(* IEC 61131-3 sources: llm-plc-st-eval/data/processed_definitivo/gpt-4o-2024-08-06/C4/zero_shot, 3 files *)

(* ---- ejec_1.st ---- *)
FUNCTION_BLOCK FB_D
VAR_INPUT
    demanda : BOOL;  // Entrada que indica si hay demanda para activar las bombas.
    falla1 : BOOL;   // Entrada que indica si la bomba1 tiene una falla.
    falla2 : BOOL;   // Entrada que indica si la bomba2 tiene una falla.
END_VAR
VAR_OUTPUT
    bomba1 : BOOL;   // Salida que controla el estado de la bomba1 (activa/inactiva).
    bomba2 : BOOL;   // Salida que controla el estado de la bomba2 (activa/inactiva).
    almFalla : BOOL; // Salida que indica si hay una alarma de falla en la bomba activa.
END_VAR
VAR
    turno : BOOL;    // Variable interna que determina cuál bomba debe activarse.
    fDem : R_TRIG;   // Detector de flanco ascendente para la señal de demanda.
END_VAR

// Detecta el flanco ascendente de la señal de demanda.
fDem(CLK := demanda);

// Si se detecta un flanco ascendente en la demanda, alterna el turno.
IF fDem.Q THEN
    turno := NOT turno;
END_IF

// Si hay demanda, decide qué bomba activar según el turno y el estado de fallas.
IF demanda THEN
    IF turno THEN
        // Si es el turno de la bomba1, actívala si no hay falla.
        bomba1 := NOT falla1;
        // Activa la bomba2 solo si la bomba1 falla y la bomba2 no tiene falla.
        bomba2 := falla1 AND NOT falla2;
        // Genera alarma si la bomba1 tiene falla.
        almFalla := falla1;
    ELSE
        // Si es el turno de la bomba2, actívala si no hay falla.
        bomba2 := NOT falla2;
        // Activa la bomba1 solo si la bomba2 falla y la bomba1 no tiene falla.
        bomba1 := falla2 AND NOT falla1;
        // Genera alarma si la bomba2 tiene falla.
        almFalla := falla2;
    END_IF
ELSE
    // Si no hay demanda, ambas bombas están inactivas y no hay alarma.
    bomba1 := FALSE;
    bomba2 := FALSE;
    almFalla := FALSE;
END_IF
END_FUNCTION_BLOCK

(* ---- ejec_2.st ---- *)
FUNCTION_BLOCK FB_D
VAR_INPUT
    demanda : BOOL; // Entrada que indica si hay demanda de bombeo
    falla1 : BOOL;  // Entrada que indica si la bomba 1 ha fallado
    falla2 : BOOL;  // Entrada que indica si la bomba 2 ha fallado
END_VAR
VAR_OUTPUT
    bomba1 : BOOL;  // Salida que controla el estado de la bomba 1
    bomba2 : BOOL;  // Salida que controla el estado de la bomba 2
    almFalla : BOOL; // Salida que indica si hay una alarma de falla
END_VAR
VAR
    turno : BOOL;   // Variable interna para alternar el uso de las bombas
    fDem : R_TRIG;  // Detector de flanco ascendente para la señal de demanda
END_VAR

// Detecta un flanco ascendente en la señal de demanda
fDem(CLK := demanda);

// Si se detecta un flanco ascendente en la demanda, alterna el turno
IF fDem.Q THEN
    turno := NOT turno;
END_IF

// Si hay demanda de bombeo
IF demanda THEN
    // Si es el turno de la bomba 1
    IF turno THEN
        bomba1 := NOT falla1; // Activa la bomba 1 si no hay falla
        bomba2 := falla1 AND NOT falla2; // Activa la bomba 2 si la bomba 1 falla y la bomba 2 no
        almFalla := falla1; // Activa la alarma si la bomba 1 falla
    ELSE
        // Si es el turno de la bomba 2
        bomba2 := NOT falla2; // Activa la bomba 2 si no hay falla
        bomba1 := falla2 AND NOT falla1; // Activa la bomba 1 si la bomba 2 falla y la bomba 1 no
        almFalla := falla2; // Activa la alarma si la bomba 2 falla
    END_IF
ELSE
    // Si no hay demanda, apaga ambas bombas y resetea la alarma
    bomba1 := FALSE;
    bomba2 := FALSE;
    almFalla := FALSE;
END_IF
END_FUNCTION_BLOCK

(* ---- ejec_3.st ---- *)
FUNCTION_BLOCK FB_D
VAR_INPUT
    demanda : BOOL;  // Entrada que indica si hay demanda de bombeo.
    falla1 : BOOL;   // Entrada que indica si la bomba1 está en estado de falla.
    falla2 : BOOL;   // Entrada que indica si la bomba2 está en estado de falla.
END_VAR
VAR_OUTPUT
    bomba1 : BOOL;   // Salida que controla el estado de la bomba1.
    bomba2 : BOOL;   // Salida que controla el estado de la bomba2.
    almFalla : BOOL; // Salida que indica si hay una alarma de falla.
END_VAR
VAR
    turno : BOOL;    // Variable interna que determina el turno de operación de las bombas.
    fDem : R_TRIG;   // Detector de flanco ascendente para la señal de demanda.
END_VAR

// Detecta el flanco ascendente de la señal de demanda.
fDem(CLK := demanda);

// Si se detecta un flanco ascendente en la demanda, se alterna el turno.
IF fDem.Q THEN
    turno := NOT turno;
END_IF

// Si hay demanda de bombeo, se evalúa el turno y el estado de falla de las bombas.
IF demanda THEN
    IF turno THEN
        // Si es el turno de bomba1, se activa si no está en falla.
        bomba1 := NOT falla1;
        // Si bomba1 está en falla, se activa bomba2 si no está en falla.
        bomba2 := falla1 AND NOT falla2;
        // Se genera una alarma si bomba1 está en falla.
        almFalla := falla1;
    ELSE
        // Si es el turno de bomba2, se activa si no está en falla.
        bomba2 := NOT falla2;
        // Si bomba2 está en falla, se activa bomba1 si no está en falla.
        bomba1 := falla2 AND NOT falla1;
        // Se genera una alarma si bomba2 está en falla.
        almFalla := falla2;
    END_IF
ELSE
    // Si no hay demanda, ambas bombas están desactivadas y no hay alarma.
    bomba1 := FALSE;
    bomba2 := FALSE;
    almFalla := FALSE;
END_IF
END_FUNCTION_BLOCK
